// TIA Portal V20 export
// export: Created 2026-10-20T12:51:33.3574785Z, ExportSetting WithDefaults, DisplayName Totally Integrated Automation Portal, DisplayVersion V20 Update 6, DisplayName TIA Portal Openness, DisplayVersion V20 Update 6, DisplayName TIA Portal Version Control Interface, DisplayVersion V20 Update 6, DisplayName SINAMICS Startdrive Advanced, DisplayVersion V20 SP1, DisplayName SINAMICS Startdrive G130, G150, S120, S150, SINAMICS MV, G220, S200, S210, DisplayVersion V20 SP1, DisplayName SINAMICS Startdrive G110M, G120, G120C, G120D, G120P, G115D, DisplayVersion V20 SP1, DisplayName STEP 7 Professional, DisplayVersion V20 Update 6, DisplayName STEP 7 Safety, DisplayVersion V20 Update 2, DisplayName WinCC Basic/Comfort/Advanced, DisplayVersion V20 Update 6, DisplayName WinCC Unified, DisplayVersion V20 Update 6
FUNCTION "Bypass assignments_0" : Void   // FC34, F_LAD
{ S7_Optimized_Access := 'TRUE' }
VERSION : 0.1
// stored: AutoNumber true, IsIECCheckEnabled false, UDAEnableTagReadback false
BEGIN

REGION Network 1
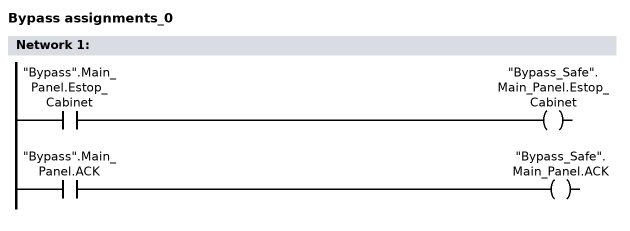
   RUNG wire#powerrail
      Contact( "Bypass".Main_Panel.Estop_Cabinet )
      Coil( "Bypass_Safe".Main_Panel.Estop_Cabinet )
   END_RUNG
   RUNG wire#powerrail
      Contact( "Bypass".Main_Panel.ACK )
      Coil( "Bypass_Safe".Main_Panel.ACK )
   END_RUNG
   // the same network as SCL:
   "Bypass_Safe".Main_Panel.Estop_Cabinet := "Bypass".Main_Panel.Estop_Cabinet;
   "Bypass_Safe".Main_Panel.ACK := "Bypass".Main_Panel.ACK;
END_REGION
END_FUNCTION
